// TIA Portal V20 export
TYPE "Schrittkettenaufruf"
   STRUCT
      OFF_SQ : Bool;
      INIT_SQ : Bool;
      ACK_EF : Bool;
      HALT_SQ : Bool;
      HALT_TM : Bool;
      ZERO_OP : Bool;
      EN_IL : Bool;
      EN_SV : Bool;
      S_PREV : Bool;
      S_NEXT : Bool;
      SW_AUTO : Bool;
      SW_TAP : Bool;
      SW_MAN : Bool;
      S_SEL : Int;
      S_ON : Bool;
      S_OFF : Bool;
      T_PUSH : Bool;
      S_NO : Int;
      S_MORE : Bool;
      S_ACTIVE : Bool;
      ERR_FLT : Bool;
      SQ_HALTED : Bool;
      TM_HALTED : Bool;
      OP_ZEROED : Bool;
      IL_ENABELD : Bool;
      SV_ENABELD : Bool;
      AUTO_ON : Bool;
      TAP_ON : Bool;
      MAN_ON : Bool;
   END_STRUCT;
END_TYPE
